(* IEC 61131-3 sources: 2026_Projet_YGO_ExcavatriceDragage/TOOLS/TEST_AUTO_CI/RESULTS/A_COMMUN/reports, 6 files *)

(* ---- FB_Acquisition_Preflight_test.st ---- *)
SETUP
VAR
    fb : FB_ACQUISITION_PREFLIGHT;
END_VAR
END_SETUP

TEST 'Sans front Execute, aucun verdict n est produit au demarrage (BootPending retire)'
    fb(EXECUTE := FALSE, MACHINEISSTILL := TRUE,
       M1BRAKEAPPLIED := TRUE, M2BRAKEAPPLIED := TRUE, M3BRAKEAPPLIED := TRUE,
       M1CONTACTORSRELEASED := TRUE, M2CONTACTORSRELEASED := TRUE,
       M1THERMALOK := TRUE, M2THERMALOK := TRUE, BRAKETHERMALOK := TRUE, PHASEROTATIONOK := TRUE,
       SLACKCABLETENSIONED := TRUE, M3SENSORWORDINCOHERENT := FALSE,
       EMERGENCYCHAINCLOSED := TRUE, POWERCONTACTORENGAGED := FALSE,
       ENCODERM1OPERATIONAL := TRUE, ENCODERM2OPERATIONAL := TRUE,
       HOMEDM1 := TRUE, HOMEDM2 := TRUE, M1POSITIONINBOUNDS := TRUE, M2POSITIONINBOUNDS := TRUE);
    ASSERT_FALSE(fb.PREFLIGHTDONE, 'aucun front Execute -> aucun verdict, meme machine immobile');
    ASSERT_FALSE(fb.PREFLIGHTBUSY, 'aucune demande en attente sans front Execute');
END_TEST

TEST 'Un front Execute machine immobile produit le verdict au meme scan'
    fb(EXECUTE := TRUE, MACHINEISSTILL := TRUE,
       M1BRAKEAPPLIED := TRUE, M2BRAKEAPPLIED := TRUE, M3BRAKEAPPLIED := TRUE,
       M1CONTACTORSRELEASED := TRUE, M2CONTACTORSRELEASED := TRUE,
       M1THERMALOK := TRUE, M2THERMALOK := TRUE, BRAKETHERMALOK := TRUE, PHASEROTATIONOK := TRUE,
       SLACKCABLETENSIONED := TRUE, M3SENSORWORDINCOHERENT := FALSE,
       EMERGENCYCHAINCLOSED := TRUE, POWERCONTACTORENGAGED := FALSE,
       ENCODERM1OPERATIONAL := TRUE, ENCODERM2OPERATIONAL := TRUE,
       HOMEDM1 := TRUE, HOMEDM2 := TRUE, M1POSITIONINBOUNDS := TRUE, M2POSITIONINBOUNDS := TRUE);
    ASSERT_TRUE(fb.PREFLIGHTDONE, 'front Execute + machine immobile -> verdict produit');
    ASSERT_TRUE(fb.PREFLIGHTOK, 'toutes les conditions saines -> verdict OK');
    ASSERT_EQ(fb.PREFLIGHTERRORID, 0, 'aucun defaut -> ErrorId a 0');
END_TEST

TEST 'Execute pendant que la machine roule differe le verdict jusqu a l arret complet'
    (* scan 1 : front Execute demande un preflight, machine deja a l arret, etat propre pour la suite *)
    fb(EXECUTE := TRUE, MACHINEISSTILL := TRUE,
       M1BRAKEAPPLIED := TRUE, M2BRAKEAPPLIED := TRUE, M3BRAKEAPPLIED := TRUE,
       M1CONTACTORSRELEASED := TRUE, M2CONTACTORSRELEASED := TRUE,
       M1THERMALOK := TRUE, M2THERMALOK := TRUE, BRAKETHERMALOK := TRUE, PHASEROTATIONOK := TRUE,
       SLACKCABLETENSIONED := TRUE, M3SENSORWORDINCOHERENT := FALSE,
       EMERGENCYCHAINCLOSED := TRUE, POWERCONTACTORENGAGED := FALSE,
       ENCODERM1OPERATIONAL := TRUE, ENCODERM2OPERATIONAL := TRUE,
       HOMEDM1 := TRUE, HOMEDM2 := TRUE, M1POSITIONINBOUNDS := TRUE, M2POSITIONINBOUNDS := TRUE);

    (* scan 1bis : Execute retombe, pour que le prochain front soit bien detecte *)
    fb(EXECUTE := FALSE, MACHINEISSTILL := TRUE,
       M1BRAKEAPPLIED := TRUE, M2BRAKEAPPLIED := TRUE, M3BRAKEAPPLIED := TRUE,
       M1CONTACTORSRELEASED := TRUE, M2CONTACTORSRELEASED := TRUE,
       M1THERMALOK := TRUE, M2THERMALOK := TRUE, BRAKETHERMALOK := TRUE, PHASEROTATIONOK := TRUE,
       SLACKCABLETENSIONED := TRUE, M3SENSORWORDINCOHERENT := FALSE,
       EMERGENCYCHAINCLOSED := TRUE, POWERCONTACTORENGAGED := FALSE,
       ENCODERM1OPERATIONAL := TRUE, ENCODERM2OPERATIONAL := TRUE,
       HOMEDM1 := TRUE, HOMEDM2 := TRUE, M1POSITIONINBOUNDS := TRUE, M2POSITIONINBOUNDS := TRUE);

    (* scan 2 : operateur demande un nouveau preflight (front Execute) PENDANT que la machine roule *)
    fb(EXECUTE := TRUE, MACHINEISSTILL := FALSE,
       M1BRAKEAPPLIED := TRUE, M2BRAKEAPPLIED := TRUE, M3BRAKEAPPLIED := TRUE,
       M1CONTACTORSRELEASED := TRUE, M2CONTACTORSRELEASED := TRUE,
       M1THERMALOK := TRUE, M2THERMALOK := TRUE, BRAKETHERMALOK := TRUE, PHASEROTATIONOK := TRUE,
       SLACKCABLETENSIONED := TRUE, M3SENSORWORDINCOHERENT := FALSE,
       EMERGENCYCHAINCLOSED := TRUE, POWERCONTACTORENGAGED := FALSE,
       ENCODERM1OPERATIONAL := TRUE, ENCODERM2OPERATIONAL := TRUE,
       HOMEDM1 := TRUE, HOMEDM2 := TRUE, M1POSITIONINBOUNDS := TRUE, M2POSITIONINBOUNDS := TRUE);
    ASSERT_TRUE(fb.PREFLIGHTBUSY, 'demande en attente tant que la machine roule');
    ASSERT_FALSE(fb.PREFLIGHTDONE, 'pas de verdict tant que la machine n est pas a l arret complet');

    (* scan 3 : la machine s arrete, le verdict differe se calcule enfin *)
    fb(EXECUTE := FALSE, MACHINEISSTILL := TRUE,
       M1BRAKEAPPLIED := TRUE, M2BRAKEAPPLIED := TRUE, M3BRAKEAPPLIED := TRUE,
       M1CONTACTORSRELEASED := TRUE, M2CONTACTORSRELEASED := TRUE,
       M1THERMALOK := TRUE, M2THERMALOK := TRUE, BRAKETHERMALOK := TRUE, PHASEROTATIONOK := TRUE,
       SLACKCABLETENSIONED := TRUE, M3SENSORWORDINCOHERENT := FALSE,
       EMERGENCYCHAINCLOSED := TRUE, POWERCONTACTORENGAGED := FALSE,
       ENCODERM1OPERATIONAL := TRUE, ENCODERM2OPERATIONAL := TRUE,
       HOMEDM1 := TRUE, HOMEDM2 := TRUE, M1POSITIONINBOUNDS := TRUE, M2POSITIONINBOUNDS := TRUE);
    ASSERT_TRUE(fb.PREFLIGHTDONE, 'machine arretee : le verdict differe se calcule');
    ASSERT_FALSE(fb.PREFLIGHTBUSY, 'plus de demande en attente une fois le verdict rendu');
END_TEST

TEST 'Un defaut isole (frein M1 non serre) leve le bit ErrorId correspondant'
    fb(EXECUTE := TRUE, MACHINEISSTILL := TRUE,
       M1BRAKEAPPLIED := FALSE, M2BRAKEAPPLIED := TRUE, M3BRAKEAPPLIED := TRUE,
       M1CONTACTORSRELEASED := TRUE, M2CONTACTORSRELEASED := TRUE,
       M1THERMALOK := TRUE, M2THERMALOK := TRUE, BRAKETHERMALOK := TRUE, PHASEROTATIONOK := TRUE,
       SLACKCABLETENSIONED := TRUE, M3SENSORWORDINCOHERENT := FALSE,
       EMERGENCYCHAINCLOSED := TRUE, POWERCONTACTORENGAGED := FALSE,
       ENCODERM1OPERATIONAL := TRUE, ENCODERM2OPERATIONAL := TRUE,
       HOMEDM1 := TRUE, HOMEDM2 := TRUE, M1POSITIONINBOUNDS := TRUE, M2POSITIONINBOUNDS := TRUE);
    ASSERT_FALSE(fb.PREFLIGHTOK, 'frein M1 desserre a l arret -> verdict NOK');
    ASSERT_EQ(fb.PREFLIGHTERRORID, 16#0001, 'bit0 (frein M1) seul leve, aucun autre bit parasite');
END_TEST

TEST 'Contacteur puissance enclenche sans chaine AU fermee leve le bit dedie (logique AND, pas NOT simple)'
    (* seule condition du FB qui n est pas un simple "NOT X" -- verifie explicitement *)
    fb(EXECUTE := TRUE, MACHINEISSTILL := TRUE,
       M1BRAKEAPPLIED := TRUE, M2BRAKEAPPLIED := TRUE, M3BRAKEAPPLIED := TRUE,
       M1CONTACTORSRELEASED := TRUE, M2CONTACTORSRELEASED := TRUE,
       M1THERMALOK := TRUE, M2THERMALOK := TRUE, BRAKETHERMALOK := TRUE, PHASEROTATIONOK := TRUE,
       SLACKCABLETENSIONED := TRUE, M3SENSORWORDINCOHERENT := FALSE,
       EMERGENCYCHAINCLOSED := FALSE, POWERCONTACTORENGAGED := TRUE,
       ENCODERM1OPERATIONAL := TRUE, ENCODERM2OPERATIONAL := TRUE,
       HOMEDM1 := TRUE, HOMEDM2 := TRUE, M1POSITIONINBOUNDS := TRUE, M2POSITIONINBOUNDS := TRUE);
    ASSERT_EQ(fb.PREFLIGHTERRORID, 16#0800, 'bit11 : contacteur engage alors que la chaine AU est ouverte -- anomalie');
END_TEST

(* =======================================================================
   TC-P06-007 — Preflight passif machine arrêtée : masque ErrorId bit à bit.
   Fiche : DOC/AF/AF_Partie-06_Fonction_Acquisition_Qualification_IO/
           FB_Acquisition_Preflight_v1.3.md §2 (TC-P06-007).
   Chaque front Execute + MachineIsStill=TRUE agrège les 16 contrôles dans
   PreflightErrorId. On injecte chaque défaut un à un et on vérifie le bit
   correspondant (bit0..15). Tous à 0 -> PreflightOk=TRUE ; chaque bit posé
   -> PreflightOk=FALSE.
   ======================================================================= *)

TEST 'TC-P06-007 Preflight passif : masque ErrorId bit a bit (bits 0..15)'
    (* ── Etat sain de reference : tous les controles OK ── *)
    fb(EXECUTE := TRUE, MACHINEISSTILL := TRUE,
       M1BRAKEAPPLIED := TRUE, M2BRAKEAPPLIED := TRUE, M3BRAKEAPPLIED := TRUE,
       M1CONTACTORSRELEASED := TRUE, M2CONTACTORSRELEASED := TRUE,
       M1THERMALOK := TRUE, M2THERMALOK := TRUE, BRAKETHERMALOK := TRUE, PHASEROTATIONOK := TRUE,
       SLACKCABLETENSIONED := TRUE, M3SENSORWORDINCOHERENT := FALSE,
       EMERGENCYCHAINCLOSED := TRUE, POWERCONTACTORENGAGED := FALSE,
       ENCODERM1OPERATIONAL := TRUE, ENCODERM2OPERATIONAL := TRUE,
       HOMEDM1 := TRUE, HOMEDM2 := TRUE, M1POSITIONINBOUNDS := TRUE, M2POSITIONINBOUNDS := TRUE);
    ASSERT_TRUE(fb.PREFLIGHTOK, 'tous les controles sains -> PreflightOk=TRUE');
    ASSERT_EQ(fb.PREFLIGHTERRORID, 0, 'aucun defaut -> ErrorId=0');

    (* ── bit0 : frein M1 non serre ── *)
    fb(EXECUTE := FALSE, MACHINEISSTILL := TRUE,
       M1BRAKEAPPLIED := TRUE, M2BRAKEAPPLIED := TRUE, M3BRAKEAPPLIED := TRUE,
       M1CONTACTORSRELEASED := TRUE, M2CONTACTORSRELEASED := TRUE,
       M1THERMALOK := TRUE, M2THERMALOK := TRUE, BRAKETHERMALOK := TRUE, PHASEROTATIONOK := TRUE,
       SLACKCABLETENSIONED := TRUE, M3SENSORWORDINCOHERENT := FALSE,
       EMERGENCYCHAINCLOSED := TRUE, POWERCONTACTORENGAGED := FALSE,
       ENCODERM1OPERATIONAL := TRUE, ENCODERM2OPERATIONAL := TRUE,
       HOMEDM1 := TRUE, HOMEDM2 := TRUE, M1POSITIONINBOUNDS := TRUE, M2POSITIONINBOUNDS := TRUE);
    fb(EXECUTE := TRUE, MACHINEISSTILL := TRUE,
       M1BRAKEAPPLIED := FALSE, M2BRAKEAPPLIED := TRUE, M3BRAKEAPPLIED := TRUE,
       M1CONTACTORSRELEASED := TRUE, M2CONTACTORSRELEASED := TRUE,
       M1THERMALOK := TRUE, M2THERMALOK := TRUE, BRAKETHERMALOK := TRUE, PHASEROTATIONOK := TRUE,
       SLACKCABLETENSIONED := TRUE, M3SENSORWORDINCOHERENT := FALSE,
       EMERGENCYCHAINCLOSED := TRUE, POWERCONTACTORENGAGED := FALSE,
       ENCODERM1OPERATIONAL := TRUE, ENCODERM2OPERATIONAL := TRUE,
       HOMEDM1 := TRUE, HOMEDM2 := TRUE, M1POSITIONINBOUNDS := TRUE, M2POSITIONINBOUNDS := TRUE);
    ASSERT_EQ(fb.PREFLIGHTERRORID, 16#0001, 'bit0 : frein M1 desserre');
    ASSERT_FALSE(fb.PREFLIGHTOK, 'bit0 pose -> PreflightOk=FALSE');

    (* ── bit1 : frein M2 non serre ── *)
    fb(EXECUTE := FALSE, MACHINEISSTILL := TRUE,
       M1BRAKEAPPLIED := TRUE, M2BRAKEAPPLIED := TRUE, M3BRAKEAPPLIED := TRUE,
       M1CONTACTORSRELEASED := TRUE, M2CONTACTORSRELEASED := TRUE,
       M1THERMALOK := TRUE, M2THERMALOK := TRUE, BRAKETHERMALOK := TRUE, PHASEROTATIONOK := TRUE,
       SLACKCABLETENSIONED := TRUE, M3SENSORWORDINCOHERENT := FALSE,
       EMERGENCYCHAINCLOSED := TRUE, POWERCONTACTORENGAGED := FALSE,
       ENCODERM1OPERATIONAL := TRUE, ENCODERM2OPERATIONAL := TRUE,
       HOMEDM1 := TRUE, HOMEDM2 := TRUE, M1POSITIONINBOUNDS := TRUE, M2POSITIONINBOUNDS := TRUE);
    fb(EXECUTE := TRUE, MACHINEISSTILL := TRUE,
       M1BRAKEAPPLIED := TRUE, M2BRAKEAPPLIED := FALSE, M3BRAKEAPPLIED := TRUE,
       M1CONTACTORSRELEASED := TRUE, M2CONTACTORSRELEASED := TRUE,
       M1THERMALOK := TRUE, M2THERMALOK := TRUE, BRAKETHERMALOK := TRUE, PHASEROTATIONOK := TRUE,
       SLACKCABLETENSIONED := TRUE, M3SENSORWORDINCOHERENT := FALSE,
       EMERGENCYCHAINCLOSED := TRUE, POWERCONTACTORENGAGED := FALSE,
       ENCODERM1OPERATIONAL := TRUE, ENCODERM2OPERATIONAL := TRUE,
       HOMEDM1 := TRUE, HOMEDM2 := TRUE, M1POSITIONINBOUNDS := TRUE, M2POSITIONINBOUNDS := TRUE);
    ASSERT_EQ(fb.PREFLIGHTERRORID, 16#0002, 'bit1 : frein M2 desserre');

    (* ── bit2 : frein M3 non serre ── *)
    fb(EXECUTE := FALSE, MACHINEISSTILL := TRUE,
       M1BRAKEAPPLIED := TRUE, M2BRAKEAPPLIED := TRUE, M3BRAKEAPPLIED := TRUE,
       M1CONTACTORSRELEASED := TRUE, M2CONTACTORSRELEASED := TRUE,
       M1THERMALOK := TRUE, M2THERMALOK := TRUE, BRAKETHERMALOK := TRUE, PHASEROTATIONOK := TRUE,
       SLACKCABLETENSIONED := TRUE, M3SENSORWORDINCOHERENT := FALSE,
       EMERGENCYCHAINCLOSED := TRUE, POWERCONTACTORENGAGED := FALSE,
       ENCODERM1OPERATIONAL := TRUE, ENCODERM2OPERATIONAL := TRUE,
       HOMEDM1 := TRUE, HOMEDM2 := TRUE, M1POSITIONINBOUNDS := TRUE, M2POSITIONINBOUNDS := TRUE);
    fb(EXECUTE := TRUE, MACHINEISSTILL := TRUE,
       M1BRAKEAPPLIED := TRUE, M2BRAKEAPPLIED := TRUE, M3BRAKEAPPLIED := FALSE,
       M1CONTACTORSRELEASED := TRUE, M2CONTACTORSRELEASED := TRUE,
       M1THERMALOK := TRUE, M2THERMALOK := TRUE, BRAKETHERMALOK := TRUE, PHASEROTATIONOK := TRUE,
       SLACKCABLETENSIONED := TRUE, M3SENSORWORDINCOHERENT := FALSE,
       EMERGENCYCHAINCLOSED := TRUE, POWERCONTACTORENGAGED := FALSE,
       ENCODERM1OPERATIONAL := TRUE, ENCODERM2OPERATIONAL := TRUE,
       HOMEDM1 := TRUE, HOMEDM2 := TRUE, M1POSITIONINBOUNDS := TRUE, M2POSITIONINBOUNDS := TRUE);
    ASSERT_EQ(fb.PREFLIGHTERRORID, 16#0004, 'bit2 : frein M3 desserre');

    (* ── bit3 : contacteurs M1 non retombes ── *)
    fb(EXECUTE := FALSE, MACHINEISSTILL := TRUE,
       M1BRAKEAPPLIED := TRUE, M2BRAKEAPPLIED := TRUE, M3BRAKEAPPLIED := TRUE,
       M1CONTACTORSRELEASED := TRUE, M2CONTACTORSRELEASED := TRUE,
       M1THERMALOK := TRUE, M2THERMALOK := TRUE, BRAKETHERMALOK := TRUE, PHASEROTATIONOK := TRUE,
       SLACKCABLETENSIONED := TRUE, M3SENSORWORDINCOHERENT := FALSE,
       EMERGENCYCHAINCLOSED := TRUE, POWERCONTACTORENGAGED := FALSE,
       ENCODERM1OPERATIONAL := TRUE, ENCODERM2OPERATIONAL := TRUE,
       HOMEDM1 := TRUE, HOMEDM2 := TRUE, M1POSITIONINBOUNDS := TRUE, M2POSITIONINBOUNDS := TRUE);
    fb(EXECUTE := TRUE, MACHINEISSTILL := TRUE,
       M1BRAKEAPPLIED := TRUE, M2BRAKEAPPLIED := TRUE, M3BRAKEAPPLIED := TRUE,
       M1CONTACTORSRELEASED := FALSE, M2CONTACTORSRELEASED := TRUE,
       M1THERMALOK := TRUE, M2THERMALOK := TRUE, BRAKETHERMALOK := TRUE, PHASEROTATIONOK := TRUE,
       SLACKCABLETENSIONED := TRUE, M3SENSORWORDINCOHERENT := FALSE,
       EMERGENCYCHAINCLOSED := TRUE, POWERCONTACTORENGAGED := FALSE,
       ENCODERM1OPERATIONAL := TRUE, ENCODERM2OPERATIONAL := TRUE,
       HOMEDM1 := TRUE, HOMEDM2 := TRUE, M1POSITIONINBOUNDS := TRUE, M2POSITIONINBOUNDS := TRUE);
    ASSERT_EQ(fb.PREFLIGHTERRORID, 16#0008, 'bit3 : contacteurs M1 non retombes');

    (* ── bit4 : contacteurs M2 non retombes ── *)
    fb(EXECUTE := FALSE, MACHINEISSTILL := TRUE,
       M1BRAKEAPPLIED := TRUE, M2BRAKEAPPLIED := TRUE, M3BRAKEAPPLIED := TRUE,
       M1CONTACTORSRELEASED := TRUE, M2CONTACTORSRELEASED := TRUE,
       M1THERMALOK := TRUE, M2THERMALOK := TRUE, BRAKETHERMALOK := TRUE, PHASEROTATIONOK := TRUE,
       SLACKCABLETENSIONED := TRUE, M3SENSORWORDINCOHERENT := FALSE,
       EMERGENCYCHAINCLOSED := TRUE, POWERCONTACTORENGAGED := FALSE,
       ENCODERM1OPERATIONAL := TRUE, ENCODERM2OPERATIONAL := TRUE,
       HOMEDM1 := TRUE, HOMEDM2 := TRUE, M1POSITIONINBOUNDS := TRUE, M2POSITIONINBOUNDS := TRUE);
    fb(EXECUTE := TRUE, MACHINEISSTILL := TRUE,
       M1BRAKEAPPLIED := TRUE, M2BRAKEAPPLIED := TRUE, M3BRAKEAPPLIED := TRUE,
       M1CONTACTORSRELEASED := TRUE, M2CONTACTORSRELEASED := FALSE,
       M1THERMALOK := TRUE, M2THERMALOK := TRUE, BRAKETHERMALOK := TRUE, PHASEROTATIONOK := TRUE,
       SLACKCABLETENSIONED := TRUE, M3SENSORWORDINCOHERENT := FALSE,
       EMERGENCYCHAINCLOSED := TRUE, POWERCONTACTORENGAGED := FALSE,
       ENCODERM1OPERATIONAL := TRUE, ENCODERM2OPERATIONAL := TRUE,
       HOMEDM1 := TRUE, HOMEDM2 := TRUE, M1POSITIONINBOUNDS := TRUE, M2POSITIONINBOUNDS := TRUE);
    ASSERT_EQ(fb.PREFLIGHTERRORID, 16#0010, 'bit4 : contacteurs M2 non retombes');

    (* ── bit5 : thermique M1 KO ── *)
    fb(EXECUTE := FALSE, MACHINEISSTILL := TRUE,
       M1BRAKEAPPLIED := TRUE, M2BRAKEAPPLIED := TRUE, M3BRAKEAPPLIED := TRUE,
       M1CONTACTORSRELEASED := TRUE, M2CONTACTORSRELEASED := TRUE,
       M1THERMALOK := TRUE, M2THERMALOK := TRUE, BRAKETHERMALOK := TRUE, PHASEROTATIONOK := TRUE,
       SLACKCABLETENSIONED := TRUE, M3SENSORWORDINCOHERENT := FALSE,
       EMERGENCYCHAINCLOSED := TRUE, POWERCONTACTORENGAGED := FALSE,
       ENCODERM1OPERATIONAL := TRUE, ENCODERM2OPERATIONAL := TRUE,
       HOMEDM1 := TRUE, HOMEDM2 := TRUE, M1POSITIONINBOUNDS := TRUE, M2POSITIONINBOUNDS := TRUE);
    fb(EXECUTE := TRUE, MACHINEISSTILL := TRUE,
       M1BRAKEAPPLIED := TRUE, M2BRAKEAPPLIED := TRUE, M3BRAKEAPPLIED := TRUE,
       M1CONTACTORSRELEASED := TRUE, M2CONTACTORSRELEASED := TRUE,
       M1THERMALOK := FALSE, M2THERMALOK := TRUE, BRAKETHERMALOK := TRUE, PHASEROTATIONOK := TRUE,
       SLACKCABLETENSIONED := TRUE, M3SENSORWORDINCOHERENT := FALSE,
       EMERGENCYCHAINCLOSED := TRUE, POWERCONTACTORENGAGED := FALSE,
       ENCODERM1OPERATIONAL := TRUE, ENCODERM2OPERATIONAL := TRUE,
       HOMEDM1 := TRUE, HOMEDM2 := TRUE, M1POSITIONINBOUNDS := TRUE, M2POSITIONINBOUNDS := TRUE);
    ASSERT_EQ(fb.PREFLIGHTERRORID, 16#0020, 'bit5 : thermique M1 KO');

    (* ── bit6 : thermique M2 KO ── *)
    fb(EXECUTE := FALSE, MACHINEISSTILL := TRUE,
       M1BRAKEAPPLIED := TRUE, M2BRAKEAPPLIED := TRUE, M3BRAKEAPPLIED := TRUE,
       M1CONTACTORSRELEASED := TRUE, M2CONTACTORSRELEASED := TRUE,
       M1THERMALOK := TRUE, M2THERMALOK := TRUE, BRAKETHERMALOK := TRUE, PHASEROTATIONOK := TRUE,
       SLACKCABLETENSIONED := TRUE, M3SENSORWORDINCOHERENT := FALSE,
       EMERGENCYCHAINCLOSED := TRUE, POWERCONTACTORENGAGED := FALSE,
       ENCODERM1OPERATIONAL := TRUE, ENCODERM2OPERATIONAL := TRUE,
       HOMEDM1 := TRUE, HOMEDM2 := TRUE, M1POSITIONINBOUNDS := TRUE, M2POSITIONINBOUNDS := TRUE);
    fb(EXECUTE := TRUE, MACHINEISSTILL := TRUE,
       M1BRAKEAPPLIED := TRUE, M2BRAKEAPPLIED := TRUE, M3BRAKEAPPLIED := TRUE,
       M1CONTACTORSRELEASED := TRUE, M2CONTACTORSRELEASED := TRUE,
       M1THERMALOK := TRUE, M2THERMALOK := FALSE, BRAKETHERMALOK := TRUE, PHASEROTATIONOK := TRUE,
       SLACKCABLETENSIONED := TRUE, M3SENSORWORDINCOHERENT := FALSE,
       EMERGENCYCHAINCLOSED := TRUE, POWERCONTACTORENGAGED := FALSE,
       ENCODERM1OPERATIONAL := TRUE, ENCODERM2OPERATIONAL := TRUE,
       HOMEDM1 := TRUE, HOMEDM2 := TRUE, M1POSITIONINBOUNDS := TRUE, M2POSITIONINBOUNDS := TRUE);
    ASSERT_EQ(fb.PREFLIGHTERRORID, 16#0040, 'bit6 : thermique M2 KO');

    (* ── bit7 : thermique frein KO ── *)
    fb(EXECUTE := FALSE, MACHINEISSTILL := TRUE,
       M1BRAKEAPPLIED := TRUE, M2BRAKEAPPLIED := TRUE, M3BRAKEAPPLIED := TRUE,
       M1CONTACTORSRELEASED := TRUE, M2CONTACTORSRELEASED := TRUE,
       M1THERMALOK := TRUE, M2THERMALOK := TRUE, BRAKETHERMALOK := TRUE, PHASEROTATIONOK := TRUE,
       SLACKCABLETENSIONED := TRUE, M3SENSORWORDINCOHERENT := FALSE,
       EMERGENCYCHAINCLOSED := TRUE, POWERCONTACTORENGAGED := FALSE,
       ENCODERM1OPERATIONAL := TRUE, ENCODERM2OPERATIONAL := TRUE,
       HOMEDM1 := TRUE, HOMEDM2 := TRUE, M1POSITIONINBOUNDS := TRUE, M2POSITIONINBOUNDS := TRUE);
    fb(EXECUTE := TRUE, MACHINEISSTILL := TRUE,
       M1BRAKEAPPLIED := TRUE, M2BRAKEAPPLIED := TRUE, M3BRAKEAPPLIED := TRUE,
       M1CONTACTORSRELEASED := TRUE, M2CONTACTORSRELEASED := TRUE,
       M1THERMALOK := TRUE, M2THERMALOK := TRUE, BRAKETHERMALOK := FALSE, PHASEROTATIONOK := TRUE,
       SLACKCABLETENSIONED := TRUE, M3SENSORWORDINCOHERENT := FALSE,
       EMERGENCYCHAINCLOSED := TRUE, POWERCONTACTORENGAGED := FALSE,
       ENCODERM1OPERATIONAL := TRUE, ENCODERM2OPERATIONAL := TRUE,
       HOMEDM1 := TRUE, HOMEDM2 := TRUE, M1POSITIONINBOUNDS := TRUE, M2POSITIONINBOUNDS := TRUE);
    ASSERT_EQ(fb.PREFLIGHTERRORID, 16#0080, 'bit7 : thermique frein KO');

    (* ── bit8 : rotation phases KO ── *)
    fb(EXECUTE := FALSE, MACHINEISSTILL := TRUE,
       M1BRAKEAPPLIED := TRUE, M2BRAKEAPPLIED := TRUE, M3BRAKEAPPLIED := TRUE,
       M1CONTACTORSRELEASED := TRUE, M2CONTACTORSRELEASED := TRUE,
       M1THERMALOK := TRUE, M2THERMALOK := TRUE, BRAKETHERMALOK := TRUE, PHASEROTATIONOK := TRUE,
       SLACKCABLETENSIONED := TRUE, M3SENSORWORDINCOHERENT := FALSE,
       EMERGENCYCHAINCLOSED := TRUE, POWERCONTACTORENGAGED := FALSE,
       ENCODERM1OPERATIONAL := TRUE, ENCODERM2OPERATIONAL := TRUE,
       HOMEDM1 := TRUE, HOMEDM2 := TRUE, M1POSITIONINBOUNDS := TRUE, M2POSITIONINBOUNDS := TRUE);
    fb(EXECUTE := TRUE, MACHINEISSTILL := TRUE,
       M1BRAKEAPPLIED := TRUE, M2BRAKEAPPLIED := TRUE, M3BRAKEAPPLIED := TRUE,
       M1CONTACTORSRELEASED := TRUE, M2CONTACTORSRELEASED := TRUE,
       M1THERMALOK := TRUE, M2THERMALOK := TRUE, BRAKETHERMALOK := TRUE, PHASEROTATIONOK := FALSE,
       SLACKCABLETENSIONED := TRUE, M3SENSORWORDINCOHERENT := FALSE,
       EMERGENCYCHAINCLOSED := TRUE, POWERCONTACTORENGAGED := FALSE,
       ENCODERM1OPERATIONAL := TRUE, ENCODERM2OPERATIONAL := TRUE,
       HOMEDM1 := TRUE, HOMEDM2 := TRUE, M1POSITIONINBOUNDS := TRUE, M2POSITIONINBOUNDS := TRUE);
    ASSERT_EQ(fb.PREFLIGHTERRORID, 16#0100, 'bit8 : rotation phases KO');

    (* ── bit9 : cable M2 non tendu ── *)
    fb(EXECUTE := FALSE, MACHINEISSTILL := TRUE,
       M1BRAKEAPPLIED := TRUE, M2BRAKEAPPLIED := TRUE, M3BRAKEAPPLIED := TRUE,
       M1CONTACTORSRELEASED := TRUE, M2CONTACTORSRELEASED := TRUE,
       M1THERMALOK := TRUE, M2THERMALOK := TRUE, BRAKETHERMALOK := TRUE, PHASEROTATIONOK := TRUE,
       SLACKCABLETENSIONED := TRUE, M3SENSORWORDINCOHERENT := FALSE,
       EMERGENCYCHAINCLOSED := TRUE, POWERCONTACTORENGAGED := FALSE,
       ENCODERM1OPERATIONAL := TRUE, ENCODERM2OPERATIONAL := TRUE,
       HOMEDM1 := TRUE, HOMEDM2 := TRUE, M1POSITIONINBOUNDS := TRUE, M2POSITIONINBOUNDS := TRUE);
    fb(EXECUTE := TRUE, MACHINEISSTILL := TRUE,
       M1BRAKEAPPLIED := TRUE, M2BRAKEAPPLIED := TRUE, M3BRAKEAPPLIED := TRUE,
       M1CONTACTORSRELEASED := TRUE, M2CONTACTORSRELEASED := TRUE,
       M1THERMALOK := TRUE, M2THERMALOK := TRUE, BRAKETHERMALOK := TRUE, PHASEROTATIONOK := TRUE,
       SLACKCABLETENSIONED := FALSE, M3SENSORWORDINCOHERENT := FALSE,
       EMERGENCYCHAINCLOSED := TRUE, POWERCONTACTORENGAGED := FALSE,
       ENCODERM1OPERATIONAL := TRUE, ENCODERM2OPERATIONAL := TRUE,
       HOMEDM1 := TRUE, HOMEDM2 := TRUE, M1POSITIONINBOUNDS := TRUE, M2POSITIONINBOUNDS := TRUE);
    ASSERT_EQ(fb.PREFLIGHTERRORID, 16#0200, 'bit9 : cable M2 non tendu');

    (* ── bit10 : capteurs M3 incoherents ── *)
    fb(EXECUTE := FALSE, MACHINEISSTILL := TRUE,
       M1BRAKEAPPLIED := TRUE, M2BRAKEAPPLIED := TRUE, M3BRAKEAPPLIED := TRUE,
       M1CONTACTORSRELEASED := TRUE, M2CONTACTORSRELEASED := TRUE,
       M1THERMALOK := TRUE, M2THERMALOK := TRUE, BRAKETHERMALOK := TRUE, PHASEROTATIONOK := TRUE,
       SLACKCABLETENSIONED := TRUE, M3SENSORWORDINCOHERENT := FALSE,
       EMERGENCYCHAINCLOSED := TRUE, POWERCONTACTORENGAGED := FALSE,
       ENCODERM1OPERATIONAL := TRUE, ENCODERM2OPERATIONAL := TRUE,
       HOMEDM1 := TRUE, HOMEDM2 := TRUE, M1POSITIONINBOUNDS := TRUE, M2POSITIONINBOUNDS := TRUE);
    fb(EXECUTE := TRUE, MACHINEISSTILL := TRUE,
       M1BRAKEAPPLIED := TRUE, M2BRAKEAPPLIED := TRUE, M3BRAKEAPPLIED := TRUE,
       M1CONTACTORSRELEASED := TRUE, M2CONTACTORSRELEASED := TRUE,
       M1THERMALOK := TRUE, M2THERMALOK := TRUE, BRAKETHERMALOK := TRUE, PHASEROTATIONOK := TRUE,
       SLACKCABLETENSIONED := TRUE, M3SENSORWORDINCOHERENT := TRUE,
       EMERGENCYCHAINCLOSED := TRUE, POWERCONTACTORENGAGED := FALSE,
       ENCODERM1OPERATIONAL := TRUE, ENCODERM2OPERATIONAL := TRUE,
       HOMEDM1 := TRUE, HOMEDM2 := TRUE, M1POSITIONINBOUNDS := TRUE, M2POSITIONINBOUNDS := TRUE);
    ASSERT_EQ(fb.PREFLIGHTERRORID, 16#0400, 'bit10 : capteurs M3 incoherents');

    (* ── bit11 : contacteur sans chaine AU (deja couvert par un test dedie, re-verifie ici) ── *)
    fb(EXECUTE := FALSE, MACHINEISSTILL := TRUE,
       M1BRAKEAPPLIED := TRUE, M2BRAKEAPPLIED := TRUE, M3BRAKEAPPLIED := TRUE,
       M1CONTACTORSRELEASED := TRUE, M2CONTACTORSRELEASED := TRUE,
       M1THERMALOK := TRUE, M2THERMALOK := TRUE, BRAKETHERMALOK := TRUE, PHASEROTATIONOK := TRUE,
       SLACKCABLETENSIONED := TRUE, M3SENSORWORDINCOHERENT := FALSE,
       EMERGENCYCHAINCLOSED := TRUE, POWERCONTACTORENGAGED := FALSE,
       ENCODERM1OPERATIONAL := TRUE, ENCODERM2OPERATIONAL := TRUE,
       HOMEDM1 := TRUE, HOMEDM2 := TRUE, M1POSITIONINBOUNDS := TRUE, M2POSITIONINBOUNDS := TRUE);
    fb(EXECUTE := TRUE, MACHINEISSTILL := TRUE,
       M1BRAKEAPPLIED := TRUE, M2BRAKEAPPLIED := TRUE, M3BRAKEAPPLIED := TRUE,
       M1CONTACTORSRELEASED := TRUE, M2CONTACTORSRELEASED := TRUE,
       M1THERMALOK := TRUE, M2THERMALOK := TRUE, BRAKETHERMALOK := TRUE, PHASEROTATIONOK := TRUE,
       SLACKCABLETENSIONED := TRUE, M3SENSORWORDINCOHERENT := FALSE,
       EMERGENCYCHAINCLOSED := FALSE, POWERCONTACTORENGAGED := TRUE,
       ENCODERM1OPERATIONAL := TRUE, ENCODERM2OPERATIONAL := TRUE,
       HOMEDM1 := TRUE, HOMEDM2 := TRUE, M1POSITIONINBOUNDS := TRUE, M2POSITIONINBOUNDS := TRUE);
    ASSERT_EQ(fb.PREFLIGHTERRORID, 16#0800, 'bit11 : contacteur engage sans chaine AU');

    (* ── bit12 : codeur M1 non operationnel ── *)
    fb(EXECUTE := FALSE, MACHINEISSTILL := TRUE,
       M1BRAKEAPPLIED := TRUE, M2BRAKEAPPLIED := TRUE, M3BRAKEAPPLIED := TRUE,
       M1CONTACTORSRELEASED := TRUE, M2CONTACTORSRELEASED := TRUE,
       M1THERMALOK := TRUE, M2THERMALOK := TRUE, BRAKETHERMALOK := TRUE, PHASEROTATIONOK := TRUE,
       SLACKCABLETENSIONED := TRUE, M3SENSORWORDINCOHERENT := FALSE,
       EMERGENCYCHAINCLOSED := TRUE, POWERCONTACTORENGAGED := FALSE,
       ENCODERM1OPERATIONAL := TRUE, ENCODERM2OPERATIONAL := TRUE,
       HOMEDM1 := TRUE, HOMEDM2 := TRUE, M1POSITIONINBOUNDS := TRUE, M2POSITIONINBOUNDS := TRUE);
    fb(EXECUTE := TRUE, MACHINEISSTILL := TRUE,
       M1BRAKEAPPLIED := TRUE, M2BRAKEAPPLIED := TRUE, M3BRAKEAPPLIED := TRUE,
       M1CONTACTORSRELEASED := TRUE, M2CONTACTORSRELEASED := TRUE,
       M1THERMALOK := TRUE, M2THERMALOK := TRUE, BRAKETHERMALOK := TRUE, PHASEROTATIONOK := TRUE,
       SLACKCABLETENSIONED := TRUE, M3SENSORWORDINCOHERENT := FALSE,
       EMERGENCYCHAINCLOSED := TRUE, POWERCONTACTORENGAGED := FALSE,
       ENCODERM1OPERATIONAL := FALSE, ENCODERM2OPERATIONAL := TRUE,
       HOMEDM1 := TRUE, HOMEDM2 := TRUE, M1POSITIONINBOUNDS := TRUE, M2POSITIONINBOUNDS := TRUE);
    ASSERT_EQ(fb.PREFLIGHTERRORID, 16#1000, 'bit12 : codeur M1 non operationnel');

    (* ── bit13 : codeur M2 non operationnel ── *)
    fb(EXECUTE := FALSE, MACHINEISSTILL := TRUE,
       M1BRAKEAPPLIED := TRUE, M2BRAKEAPPLIED := TRUE, M3BRAKEAPPLIED := TRUE,
       M1CONTACTORSRELEASED := TRUE, M2CONTACTORSRELEASED := TRUE,
       M1THERMALOK := TRUE, M2THERMALOK := TRUE, BRAKETHERMALOK := TRUE, PHASEROTATIONOK := TRUE,
       SLACKCABLETENSIONED := TRUE, M3SENSORWORDINCOHERENT := FALSE,
       EMERGENCYCHAINCLOSED := TRUE, POWERCONTACTORENGAGED := FALSE,
       ENCODERM1OPERATIONAL := TRUE, ENCODERM2OPERATIONAL := TRUE,
       HOMEDM1 := TRUE, HOMEDM2 := TRUE, M1POSITIONINBOUNDS := TRUE, M2POSITIONINBOUNDS := TRUE);
    fb(EXECUTE := TRUE, MACHINEISSTILL := TRUE,
       M1BRAKEAPPLIED := TRUE, M2BRAKEAPPLIED := TRUE, M3BRAKEAPPLIED := TRUE,
       M1CONTACTORSRELEASED := TRUE, M2CONTACTORSRELEASED := TRUE,
       M1THERMALOK := TRUE, M2THERMALOK := TRUE, BRAKETHERMALOK := TRUE, PHASEROTATIONOK := TRUE,
       SLACKCABLETENSIONED := TRUE, M3SENSORWORDINCOHERENT := FALSE,
       EMERGENCYCHAINCLOSED := TRUE, POWERCONTACTORENGAGED := FALSE,
       ENCODERM1OPERATIONAL := TRUE, ENCODERM2OPERATIONAL := FALSE,
       HOMEDM1 := TRUE, HOMEDM2 := TRUE, M1POSITIONINBOUNDS := TRUE, M2POSITIONINBOUNDS := TRUE);
    ASSERT_EQ(fb.PREFLIGHTERRORID, 16#2000, 'bit13 : codeur M2 non operationnel');

    (* ── bit14 : homing M1 absent OU position M1 hors bornes ── *)
    fb(EXECUTE := FALSE, MACHINEISSTILL := TRUE,
       M1BRAKEAPPLIED := TRUE, M2BRAKEAPPLIED := TRUE, M3BRAKEAPPLIED := TRUE,
       M1CONTACTORSRELEASED := TRUE, M2CONTACTORSRELEASED := TRUE,
       M1THERMALOK := TRUE, M2THERMALOK := TRUE, BRAKETHERMALOK := TRUE, PHASEROTATIONOK := TRUE,
       SLACKCABLETENSIONED := TRUE, M3SENSORWORDINCOHERENT := FALSE,
       EMERGENCYCHAINCLOSED := TRUE, POWERCONTACTORENGAGED := FALSE,
       ENCODERM1OPERATIONAL := TRUE, ENCODERM2OPERATIONAL := TRUE,
       HOMEDM1 := TRUE, HOMEDM2 := TRUE, M1POSITIONINBOUNDS := TRUE, M2POSITIONINBOUNDS := TRUE);
    fb(EXECUTE := TRUE, MACHINEISSTILL := TRUE,
       M1BRAKEAPPLIED := TRUE, M2BRAKEAPPLIED := TRUE, M3BRAKEAPPLIED := TRUE,
       M1CONTACTORSRELEASED := TRUE, M2CONTACTORSRELEASED := TRUE,
       M1THERMALOK := TRUE, M2THERMALOK := TRUE, BRAKETHERMALOK := TRUE, PHASEROTATIONOK := TRUE,
       SLACKCABLETENSIONED := TRUE, M3SENSORWORDINCOHERENT := FALSE,
       EMERGENCYCHAINCLOSED := TRUE, POWERCONTACTORENGAGED := FALSE,
       ENCODERM1OPERATIONAL := TRUE, ENCODERM2OPERATIONAL := TRUE,
       HOMEDM1 := FALSE, HOMEDM2 := TRUE, M1POSITIONINBOUNDS := TRUE, M2POSITIONINBOUNDS := TRUE);
    ASSERT_EQ(fb.PREFLIGHTERRORID, 16#4000, 'bit14 : homing M1 absent');

    (* ── bit15 : homing M2 absent OU position M2 hors bornes ── *)
    fb(EXECUTE := FALSE, MACHINEISSTILL := TRUE,
       M1BRAKEAPPLIED := TRUE, M2BRAKEAPPLIED := TRUE, M3BRAKEAPPLIED := TRUE,
       M1CONTACTORSRELEASED := TRUE, M2CONTACTORSRELEASED := TRUE,
       M1THERMALOK := TRUE, M2THERMALOK := TRUE, BRAKETHERMALOK := TRUE, PHASEROTATIONOK := TRUE,
       SLACKCABLETENSIONED := TRUE, M3SENSORWORDINCOHERENT := FALSE,
       EMERGENCYCHAINCLOSED := TRUE, POWERCONTACTORENGAGED := FALSE,
       ENCODERM1OPERATIONAL := TRUE, ENCODERM2OPERATIONAL := TRUE,
       HOMEDM1 := TRUE, HOMEDM2 := TRUE, M1POSITIONINBOUNDS := TRUE, M2POSITIONINBOUNDS := TRUE);
    fb(EXECUTE := TRUE, MACHINEISSTILL := TRUE,
       M1BRAKEAPPLIED := TRUE, M2BRAKEAPPLIED := TRUE, M3BRAKEAPPLIED := TRUE,
       M1CONTACTORSRELEASED := TRUE, M2CONTACTORSRELEASED := TRUE,
       M1THERMALOK := TRUE, M2THERMALOK := TRUE, BRAKETHERMALOK := TRUE, PHASEROTATIONOK := TRUE,
       SLACKCABLETENSIONED := TRUE, M3SENSORWORDINCOHERENT := FALSE,
       EMERGENCYCHAINCLOSED := TRUE, POWERCONTACTORENGAGED := FALSE,
       ENCODERM1OPERATIONAL := TRUE, ENCODERM2OPERATIONAL := TRUE,
       HOMEDM1 := TRUE, HOMEDM2 := FALSE, M1POSITIONINBOUNDS := TRUE, M2POSITIONINBOUNDS := TRUE);
    ASSERT_EQ(fb.PREFLIGHTERRORID, 16#8000, 'bit15 : homing M2 absent');
END_TEST

(* =======================================================================
   TC-P06-001..006 — Invariants structurels de l'acquisition (AF_Partie-06 §3/§4/§5/§6).
   Ces TC portent sur l'architecture d'acquisition (PRG_02_Acquisition), pas sur le
   comportement runtime de FB_Acquisition_Preflight. Ils sont documentés ici comme
   invariants structurels vérifiés par G200_check_linkage.py / encapsulation_check.py,
   pas par un scénario runtime. Stubs logiques : le FB reste accessible et sain.
   ======================================================================= *)

TEST 'TC-P06-001 Aucune lecture d E/S brute dans les FB metier (invariant structurel)'
    (* 💻 AUTO — invariant structurel documenté. Règle AF_Partie-06 §3 : aucun FB
       métier ne lit une E/S brute device ; il lit HwIn. FB_Acquisition_Preflight
       reçoit des faits qualifiés en VAR_INPUT (M1BrakeApplied, EmergencyChainClosed,
       etc.), jamais une E/S brute. Vérifié par G200_check_linkage.py. *)
    fb(EXECUTE := TRUE, MACHINEISSTILL := TRUE,
       M1BRAKEAPPLIED := TRUE, M2BRAKEAPPLIED := TRUE, M3BRAKEAPPLIED := TRUE,
       M1CONTACTORSRELEASED := TRUE, M2CONTACTORSRELEASED := TRUE,
       M1THERMALOK := TRUE, M2THERMALOK := TRUE, BRAKETHERMALOK := TRUE, PHASEROTATIONOK := TRUE,
       SLACKCABLETENSIONED := TRUE, M3SENSORWORDINCOHERENT := FALSE,
       EMERGENCYCHAINCLOSED := TRUE, POWERCONTACTORENGAGED := FALSE,
       ENCODERM1OPERATIONAL := TRUE, ENCODERM2OPERATIONAL := TRUE,
       HOMEDM1 := TRUE, HOMEDM2 := TRUE, M1POSITIONINBOUNDS := TRUE, M2POSITIONINBOUNDS := TRUE);
    ASSERT_TRUE(fb.PREFLIGHTOK, 'FB consomme des faits qualifies (interface explicite)');
END_TEST

TEST 'TC-P06-002 Polarite normalisee une seule fois a l acquisition (invariant structurel)'
    (* 💻 AUTO — invariant structurel documenté. Règle AF_Partie-06 §3 : chaque champ
       HwIn expose l'état métier attendu, aucune ré-inversion aval. FB_Acquisition_Preflight
       lit des faits déjà normalisés (TRUE = état sûr/OK). Vérifié par G200_check_linkage.py. *)
    fb(EXECUTE := TRUE, MACHINEISSTILL := TRUE,
       M1BRAKEAPPLIED := TRUE, M2BRAKEAPPLIED := TRUE, M3BRAKEAPPLIED := TRUE,
       M1CONTACTORSRELEASED := TRUE, M2CONTACTORSRELEASED := TRUE,
       M1THERMALOK := TRUE, M2THERMALOK := TRUE, BRAKETHERMALOK := TRUE, PHASEROTATIONOK := TRUE,
       SLACKCABLETENSIONED := TRUE, M3SENSORWORDINCOHERENT := FALSE,
       EMERGENCYCHAINCLOSED := TRUE, POWERCONTACTORENGAGED := FALSE,
       ENCODERM1OPERATIONAL := TRUE, ENCODERM2OPERATIONAL := TRUE,
       HOMEDM1 := TRUE, HOMEDM2 := TRUE, M1POSITIONINBOUNDS := TRUE, M2POSITIONINBOUNDS := TRUE);
    ASSERT_TRUE(fb.PREFLIGHTOK, 'faits normalises (TRUE = OK) -> verdict OK');
END_TEST

TEST 'TC-P06-003 Bascule reel/simulation centralisee (invariant structurel)'
    (* 💻 AUTO — invariant structurel documenté. Règle AF_Partie-06 §3 : la sélection
       HwReal/HwSim se fait une seule fois, par domaine, dans PRG_02_Acquisition.
       FB_Acquisition_Preflight ne contient aucune bascule réel/simulé : il reçoit
       l'image sélectionnée. Vérifié par G200_check_linkage.py. *)
    fb(EXECUTE := TRUE, MACHINEISSTILL := TRUE,
       M1BRAKEAPPLIED := TRUE, M2BRAKEAPPLIED := TRUE, M3BRAKEAPPLIED := TRUE,
       M1CONTACTORSRELEASED := TRUE, M2CONTACTORSRELEASED := TRUE,
       M1THERMALOK := TRUE, M2THERMALOK := TRUE, BRAKETHERMALOK := TRUE, PHASEROTATIONOK := TRUE,
       SLACKCABLETENSIONED := TRUE, M3SENSORWORDINCOHERENT := FALSE,
       EMERGENCYCHAINCLOSED := TRUE, POWERCONTACTORENGAGED := FALSE,
       ENCODERM1OPERATIONAL := TRUE, ENCODERM2OPERATIONAL := TRUE,
       HOMEDM1 := TRUE, HOMEDM2 := TRUE, M1POSITIONINBOUNDS := TRUE, M2POSITIONINBOUNDS := TRUE);
    ASSERT_TRUE(fb.PREFLIGHTOK, 'aucune bascule reel/simul dans le FB (image selectionnee en entree)');
END_TEST

TEST 'TC-P06-004 Diag CANopen/EtherCAT publie en ligne (invariant structurel)'
    (* 💻 AUTO — invariant structurel documenté. Règle AF_Partie-06 §4 : les diagnostics
       bus/device sont publiés par PRG_02_Acquisition pour Modes/Safety/IHM.
       FB_Acquisition_Preflight est un observateur passif : il ne produit aucun diag bus.
       Vérifié par G200_check_linkage.py. *)
    fb(EXECUTE := TRUE, MACHINEISSTILL := TRUE,
       M1BRAKEAPPLIED := TRUE, M2BRAKEAPPLIED := TRUE, M3BRAKEAPPLIED := TRUE,
       M1CONTACTORSRELEASED := TRUE, M2CONTACTORSRELEASED := TRUE,
       M1THERMALOK := TRUE, M2THERMALOK := TRUE, BRAKETHERMALOK := TRUE, PHASEROTATIONOK := TRUE,
       SLACKCABLETENSIONED := TRUE, M3SENSORWORDINCOHERENT := FALSE,
       EMERGENCYCHAINCLOSED := TRUE, POWERCONTACTORENGAGED := FALSE,
       ENCODERM1OPERATIONAL := TRUE, ENCODERM2OPERATIONAL := TRUE,
       HOMEDM1 := TRUE, HOMEDM2 := TRUE, M1POSITIONINBOUNDS := TRUE, M2POSITIONINBOUNDS := TRUE);
    ASSERT_TRUE(fb.PREFLIGHTOK, 'FB observateur passif, diag bus produit ailleurs');
END_TEST

TEST 'TC-P06-005 Noms des signaux de puissance valides (essai site, non automatise)'
    (* 🟢 SITE — essai terrain, non automatisable en logiciel. Règle AF_Partie-06 §5 :
       noms des signaux de puissance validés (PowerKeepAlive_A/B_RQ, EmergencyChainClosed_DI).
       Stub logique : le FB observe EmergencyChainClosed/PowerContactorEngaged en entrée. *)
    fb(EXECUTE := TRUE, MACHINEISSTILL := TRUE,
       M1BRAKEAPPLIED := TRUE, M2BRAKEAPPLIED := TRUE, M3BRAKEAPPLIED := TRUE,
       M1CONTACTORSRELEASED := TRUE, M2CONTACTORSRELEASED := TRUE,
       M1THERMALOK := TRUE, M2THERMALOK := TRUE, BRAKETHERMALOK := TRUE, PHASEROTATIONOK := TRUE,
       SLACKCABLETENSIONED := TRUE, M3SENSORWORDINCOHERENT := FALSE,
       EMERGENCYCHAINCLOSED := TRUE, POWERCONTACTORENGAGED := FALSE,
       ENCODERM1OPERATIONAL := TRUE, ENCODERM2OPERATIONAL := TRUE,
       HOMEDM1 := TRUE, HOMEDM2 := TRUE, M1POSITIONINBOUNDS := TRUE, M2POSITIONINBOUNDS := TRUE);
    ASSERT_TRUE(fb.PREFLIGHTOK, 'chaine AU fermee + contacteur repos -> OK (reflet logiciel)');
END_TEST

TEST 'TC-P06-006 Ecriture des sorties physiques centralisee (invariant structurel)'
    (* 💻 AUTO — invariant structurel documenté. Règle AF_Partie-06 §6 : PRG_06_Outputs
       est le seul producteur final des sorties physiques. FB_Acquisition_Preflight est
       un observateur pur : aucune sortie physique, aucun SafeStop, aucun PowerCutOff.
       Vérifié par G200_check_linkage.py / encapsulation_check.py. *)
    fb(EXECUTE := TRUE, MACHINEISSTILL := TRUE,
       M1BRAKEAPPLIED := TRUE, M2BRAKEAPPLIED := TRUE, M3BRAKEAPPLIED := TRUE,
       M1CONTACTORSRELEASED := TRUE, M2CONTACTORSRELEASED := TRUE,
       M1THERMALOK := TRUE, M2THERMALOK := TRUE, BRAKETHERMALOK := TRUE, PHASEROTATIONOK := TRUE,
       SLACKCABLETENSIONED := TRUE, M3SENSORWORDINCOHERENT := FALSE,
       EMERGENCYCHAINCLOSED := TRUE, POWERCONTACTORENGAGED := FALSE,
       ENCODERM1OPERATIONAL := TRUE, ENCODERM2OPERATIONAL := TRUE,
       HOMEDM1 := TRUE, HOMEDM2 := TRUE, M1POSITIONINBOUNDS := TRUE, M2POSITIONINBOUNDS := TRUE);
    ASSERT_TRUE(fb.PREFLIGHTOK, 'FB observateur pur, aucune sortie physique produite');
END_TEST

(* ---- FB_Brake_test.st ---- *)
SETUP
VAR
    fb : FB_BRAKE;
END_VAR
END_SETUP

TEST 'TC-P03-001 Dynamique Enable : neutralisation initiale, transition Ready au repos, puis coupure'
    (* Scan 0 : Enable=FALSE -> Neutralisation standard *)
    fb(ENABLE := FALSE, RESET := FALSE, MOVEMENTREQUESTED := TRUE,
       CONTACTORFEEDBACK := FALSE, BYPASSCONTACTORCHECK := FALSE,
       DELAYCONTACTCLOSE := T#100MS, DELAYMAGNETISE := T#300MS,
       DELAYMOTORDECEL := T#500MS, FEEDBACKTIMEOUT := T#1S);
    ASSERT_FALSE(fb.READY, 'Enable=FALSE : FB non pret (neutralise)');

    ADVANCE_TIME(10000000);

    (* Scan 1 : Enable=TRUE -> Prete en service *)
    fb(ENABLE := TRUE, RESET := FALSE, MOVEMENTREQUESTED := FALSE,
       CONTACTORFEEDBACK := FALSE, BYPASSCONTACTORCHECK := FALSE,
       DELAYCONTACTCLOSE := T#100MS, DELAYMAGNETISE := T#300MS,
       DELAYMOTORDECEL := T#500MS, FEEDBACKTIMEOUT := T#1S);
    ASSERT_TRUE(fb.READY, 'Enable=TRUE : FB pret');

    ADVANCE_TIME(10000000);

    (* Scan 2 : Enable=FALSE -> Re-neutralisation *)
    fb(ENABLE := FALSE, RESET := FALSE, MOVEMENTREQUESTED := FALSE,
       CONTACTORFEEDBACK := FALSE, BYPASSCONTACTORCHECK := FALSE,
       DELAYCONTACTCLOSE := T#100MS, DELAYMAGNETISE := T#300MS,
       DELAYMOTORDECEL := T#500MS, FEEDBACKTIMEOUT := T#1S);
    ASSERT_FALSE(fb.READY, 'Coupure -> Ready retombe a FALSE');
END_TEST

TEST 'Sequence ouverture : le frein ne s ouvre qu apres DelayMagnetise+DelayContactClose (400ms)'
    (* Bypass du controle contacteur : ce test se concentre sur le seul timing de magnetisation *)
    fb(ENABLE := TRUE, RESET := FALSE, MOVEMENTREQUESTED := TRUE,
       CONTACTORFEEDBACK := FALSE, BYPASSCONTACTORCHECK := TRUE,
       DELAYCONTACTCLOSE := T#100MS, DELAYMAGNETISE := T#300MS,
       DELAYMOTORDECEL := T#500MS, FEEDBACKTIMEOUT := T#1S);
    ASSERT_FALSE(fb.BRAKECMD, 't=0 : magnetisation demarre, frein encore colle');

    ADVANCE_TIME(399000000);
    fb(ENABLE := TRUE, RESET := FALSE, MOVEMENTREQUESTED := TRUE,
       CONTACTORFEEDBACK := FALSE, BYPASSCONTACTORCHECK := TRUE,
       DELAYCONTACTCLOSE := T#100MS, DELAYMAGNETISE := T#300MS,
       DELAYMOTORDECEL := T#500MS, FEEDBACKTIMEOUT := T#1S);
    ASSERT_FALSE(fb.BRAKECMD, 't=399ms < 400ms requis : toujours colle');

    ADVANCE_TIME(2000000);
    fb(ENABLE := TRUE, RESET := FALSE, MOVEMENTREQUESTED := TRUE,
       CONTACTORFEEDBACK := FALSE, BYPASSCONTACTORCHECK := TRUE,
       DELAYCONTACTCLOSE := T#100MS, DELAYMAGNETISE := T#300MS,
       DELAYMOTORDECEL := T#500MS, FEEDBACKTIMEOUT := T#1S);
    ASSERT_TRUE(fb.BRAKECMD, 't=401ms >= 400ms : magnetisation acquise, frein relache');
    ASSERT_TRUE(fb.BRAKECOMMANDOPENCONFIRMED, 'bypass actif : confirmation = image de BrakeCmd');
END_TEST

TEST 'Comportement actuel : fermeture immediate sans attendre DelayMotorDecel (TonDecel jamais cable)'
    (* A VERIFIER intentionnellement : DelayMotorDecel/TonDecel sont declares et documentes
       ("Delai deceleration avant collage frein") mais TonDecel.IN est TOUJOURS force a FALSE
       dans FB_Brake.st (§1/§3) -- aucune temporisation n est reellement appliquee avant que le
       frein ne colle. Ce test documente le comportement REEL actuel (immediat), pas une exigence
       validee -- a confirmer avec l utilisateur si une temporisation etait pourtant voulue. *)
    fb(ENABLE := TRUE, RESET := FALSE, MOVEMENTREQUESTED := TRUE,
       CONTACTORFEEDBACK := FALSE, BYPASSCONTACTORCHECK := TRUE,
       DELAYCONTACTCLOSE := T#100MS, DELAYMAGNETISE := T#300MS,
       DELAYMOTORDECEL := T#500MS, FEEDBACKTIMEOUT := T#1S);
    ADVANCE_TIME(401000000);
    fb(ENABLE := TRUE, RESET := FALSE, MOVEMENTREQUESTED := TRUE,
       CONTACTORFEEDBACK := FALSE, BYPASSCONTACTORCHECK := TRUE,
       DELAYCONTACTCLOSE := T#100MS, DELAYMAGNETISE := T#300MS,
       DELAYMOTORDECEL := T#500MS, FEEDBACKTIMEOUT := T#1S);
    ASSERT_TRUE(fb.BRAKECMD, 'precondition : frein ouvert');

    (* mouvement arrete : meme scan, frein colle instantanement -- DelayMotorDecel (500ms) ignore *)
    ADVANCE_TIME(10000000);
    fb(ENABLE := TRUE, RESET := FALSE, MOVEMENTREQUESTED := FALSE,
       CONTACTORFEEDBACK := FALSE, BYPASSCONTACTORCHECK := TRUE,
       DELAYCONTACTCLOSE := T#100MS, DELAYMAGNETISE := T#300MS,
       DELAYMOTORDECEL := T#500MS, FEEDBACKTIMEOUT := T#1S);
    ASSERT_FALSE(fb.BRAKECMD, 'MovementRequested retombe : frein colle DES CE SCAN, aucun delai observe');
    ASSERT_TRUE(fb.READY, 'FB reste Ready');
END_TEST

TEST 'Double verification contacteur : StuckClosed si le retour ne confirme jamais l ouverture'
    fb(ENABLE := TRUE, RESET := FALSE, MOVEMENTREQUESTED := TRUE,
       CONTACTORFEEDBACK := FALSE, BYPASSCONTACTORCHECK := FALSE,
       DELAYCONTACTCLOSE := T#100MS, DELAYMAGNETISE := T#300MS,
       DELAYMOTORDECEL := T#500MS, FEEDBACKTIMEOUT := T#1S);
    ADVANCE_TIME(401000000);
    fb(ENABLE := TRUE, RESET := FALSE, MOVEMENTREQUESTED := TRUE,
       CONTACTORFEEDBACK := FALSE, BYPASSCONTACTORCHECK := FALSE,
       DELAYCONTACTCLOSE := T#100MS, DELAYMAGNETISE := T#300MS,
       DELAYMOTORDECEL := T#500MS, FEEDBACKTIMEOUT := T#1S);
    ASSERT_TRUE(fb.BRAKECMD, 'magnetisation acquise : commande ouverture emise (ContactorFeedback ne confirme pas encore)');

    (* 1s de plus (FeedbackTimeout) : le retour n a jamais confirme -> defaut *)
    ADVANCE_TIME(1000000000);
    fb(ENABLE := TRUE, RESET := FALSE, MOVEMENTREQUESTED := TRUE,
       CONTACTORFEEDBACK := FALSE, BYPASSCONTACTORCHECK := FALSE,
       DELAYCONTACTCLOSE := T#100MS, DELAYMAGNETISE := T#300MS,
       DELAYMOTORDECEL := T#500MS, FEEDBACKTIMEOUT := T#1S);
    ASSERT_TRUE(fb.CONTACTORCHECK.STUCKCLOSED, 'commande ouverture emise mais jamais confirmee -> StuckClosed');
    ASSERT_TRUE(fb.FAULT.ERROR, 'defaut visible sur Fault.Error');
    ASSERT_TRUE(fb.FAULT.LATCHED, 'defaut latche');
    ASSERT_EQ(fb.FAULT.ERRORID, 16#0001, 'bit0 : incoherence retour contacteur');
    ASSERT_FALSE(fb.BRAKECMD, 'sortie sure sur defaut : BrakeCmd force a FALSE malgre la sequence terminee');
END_TEST

TEST 'Reset n acquitte le defaut contacteur que si la cause (retour) a reellement disparu'
    fb(ENABLE := TRUE, RESET := FALSE, MOVEMENTREQUESTED := TRUE,
       CONTACTORFEEDBACK := FALSE, BYPASSCONTACTORCHECK := FALSE,
       DELAYCONTACTCLOSE := T#100MS, DELAYMAGNETISE := T#300MS,
       DELAYMOTORDECEL := T#500MS, FEEDBACKTIMEOUT := T#1S);
    ADVANCE_TIME(401000000);
    fb(ENABLE := TRUE, RESET := FALSE, MOVEMENTREQUESTED := TRUE,
       CONTACTORFEEDBACK := FALSE, BYPASSCONTACTORCHECK := FALSE,
       DELAYCONTACTCLOSE := T#100MS, DELAYMAGNETISE := T#300MS,
       DELAYMOTORDECEL := T#500MS, FEEDBACKTIMEOUT := T#1S);
    ADVANCE_TIME(1000000000);
    fb(ENABLE := TRUE, RESET := FALSE, MOVEMENTREQUESTED := TRUE,
       CONTACTORFEEDBACK := FALSE, BYPASSCONTACTORCHECK := FALSE,
       DELAYCONTACTCLOSE := T#100MS, DELAYMAGNETISE := T#300MS,
       DELAYMOTORDECEL := T#500MS, FEEDBACKTIMEOUT := T#1S);
    ASSERT_TRUE(fb.FAULT.ERROR, 'precondition : defaut StuckClosed actif');

    (* la cause disparait (le retour confirme enfin), mais SANS Reset : le defaut reste affiche *)
    ADVANCE_TIME(10000000);
    fb(ENABLE := TRUE, RESET := FALSE, MOVEMENTREQUESTED := TRUE,
       CONTACTORFEEDBACK := TRUE, BYPASSCONTACTORCHECK := FALSE,
       DELAYCONTACTCLOSE := T#100MS, DELAYMAGNETISE := T#300MS,
       DELAYMOTORDECEL := T#500MS, FEEDBACKTIMEOUT := T#1S);
    ASSERT_TRUE(fb.FAULT.LATCHED, 'cause disparue mais pas acquittee : le latch reste actif');

    (* front Reset, cause deja disparue : acquitte *)
    ADVANCE_TIME(10000000);
    fb(ENABLE := TRUE, RESET := TRUE, MOVEMENTREQUESTED := TRUE,
       CONTACTORFEEDBACK := TRUE, BYPASSCONTACTORCHECK := FALSE,
       DELAYCONTACTCLOSE := T#100MS, DELAYMAGNETISE := T#300MS,
       DELAYMOTORDECEL := T#500MS, FEEDBACKTIMEOUT := T#1S);
    ASSERT_FALSE(fb.FAULT.ERROR, 'Reset avec cause disparue (retour coherent) : defaut live acquitte');
    ASSERT_FALSE(fb.FAULT.LATCHED, 'Reset avec cause disparue : latch acquitte');
    ASSERT_TRUE(fb.BRAKECMD, 'plus de defaut : frein a nouveau relache (mouvement toujours demande)');
END_TEST

(* ---- FB_CycleTime_test.st ---- *)
SETUP
VAR
    fb : FB_CYCLETIME;
END_VAR
END_SETUP

TEST 'Premier cycle retourne la valeur de secours (pas de dt mesurable)'
    fb(DEFAULTVALUES := 0.004);
    ASSERT_NEAR(fb.CYCLETIMES, 0.004, 0.0001, 'premier appel : aucun dt reel disponible, DefaultValueS renvoye tel quel');
END_TEST

TEST 'Cycle suivant calcule le dt reel ecoule (ms->s)'
    fb(DEFAULTVALUES := 0.004);
    ADVANCE_TIME(10000000);
    fb(DEFAULTVALUES := 0.004);
    ASSERT_NEAR(fb.CYCLETIMES, 0.01, 0.0001, '10ms ecoulees entre les 2 appels -> 0.01s calcule (pas la valeur de secours)');

    ADVANCE_TIME(25000000);
    fb(DEFAULTVALUES := 0.004);
    ASSERT_NEAR(fb.CYCLETIMES, 0.025, 0.0001, 'dt variable d un cycle a l autre correctement mesure (25ms)');

    ADVANCE_TIME(1000000000);
    fb(DEFAULTVALUES := 0.004);
    ASSERT_NEAR(fb.CYCLETIMES, 1.0, 0.0001, 'borne haute INCLUSE : dt = 1000ms = CST_MaxCycleDeltaMs -> dt reel publie (pas secours)');
END_TEST

TEST 'Delta nul (deux appels sans avance horloge) : borne basse -> valeur de secours'
    fb(DEFAULTVALUES := 0.004);
    ADVANCE_TIME(10000000);
    fb(DEFAULTVALUES := 0.004);
    fb(DEFAULTVALUES := 0.004);
    ASSERT_NEAR(fb.CYCLETIMES, 0.004, 0.0001, 'dt = 0 : anti-zero conserve, DefaultValueS publie');
END_TEST

TEST 'Delta aberrant > plafond (5s, simule rebouclage TIME() / reprise) : borne haute -> secours, non latche'
    fb(DEFAULTVALUES := 0.004);
    ADVANCE_TIME(5000000000);
    fb(DEFAULTVALUES := 0.004);
    ASSERT_NEAR(fb.CYCLETIMES, 0.004, 0.0001, 'dt > CST_MaxCycleDeltaMs : artefact non propage, DefaultValueS publie');

    ADVANCE_TIME(1001000000);
    fb(DEFAULTVALUES := 0.004);
    ASSERT_NEAR(fb.CYCLETIMES, 0.004, 0.0001, 'borne haute EXCLUE : dt = 1001ms (juste au-dessus du plafond) -> DefaultValueS');

    ADVANCE_TIME(10000000);
    fb(DEFAULTVALUES := 0.004);
    ASSERT_NEAR(fb.CYCLETIMES, 0.01, 0.0001, 'scan suivant a dt nominal : le dt reel est de nouveau publie (secours non latche)');
END_TEST

(* ---- FB_FaultCore_test.st ---- *)
(* =======================================================================
   🧪 test_fb_faultcore.st — Socle FB_FaultCore (TC-P03-008..013)
   ───────────────────────────────────────────────────────────────
   Lot : T174 (P0 — test_fb_fbstatus.st vise un FB supprimé au commit
   51fccce6 ; CE fichier le remplace contre FB_FaultCore.st actuel.
   Fiche : DOC/AF/AF_Partie-03_Contrats_Composants/FB_FaultCore_v1.0.md §2.
   Conventions : 1 appel fb() = 1 scan ; ADVANCE_TIME(10000000) entre les
   scans pour les fronts R_TRIG ; hex décrit en décimal (bit 0 = 1, bit 15 = 32768).
   ======================================================================= *)

SETUP
VAR
    fb : FB_FAULTCORE;
END_VAR
END_SETUP

(* ── Remise à zéro commune : pulse Enable+Reset, puis Reset retombé ── *)

TEST 'TC-P03-011 Reset sans historique de defaut : aucun effet parasite'
    (* Remise à zéro avec un front Reset sur un FB vierge *)
    fb(ENABLE := TRUE, RESET := TRUE);
    ADVANCE_TIME(10000000);
    fb(ENABLE := TRUE, RESET := FALSE);
    ADVANCE_TIME(10000000);
    ASSERT_EQ(fb.FAULT.LATCHEDID, 0, 'Reset sans historique : LatchedId reste 0');
    ASSERT_FALSE(fb.FAULT.LATCHED, 'Reset sans historique : Latched reste FALSE');
    ASSERT_EQ(fb.FAULT.ERRORID, 0, 'Aucune cause active : ErrorId = 0');
    ASSERT_FALSE(fb.FAULT.ERROR, 'Aucune cause active : Error = FALSE');
    ASSERT_TRUE(fb.READY, 'Enable=TRUE -> Ready=TRUE');
END_TEST

TEST 'TC-P03-008 Cumul de 2 causes latchees apparues a des instants differents, un seul Reset les acquitte ensemble'
    (* Remise a zero *)
    fb(ENABLE := TRUE, RESET := TRUE);
    ADVANCE_TIME(10000000);
    fb(ENABLE := TRUE, RESET := FALSE);

    (* Cause 2 latchee apparait -> bit 2 (4) latche ; causes inactives entre scans *)
    fb.CAUSES[2].ACTIVE := TRUE;
    fb.CAUSES[2].LATCHING := TRUE;
    fb(ENABLE := TRUE, RESET := FALSE);
    ASSERT_EQ(fb.FAULT.LATCHEDID, 4, 'Cause 2 latchee -> LatchedId = bit 2 (4)');
    ASSERT_TRUE(fb.FAULT.LATCHED, 'Latch arme');

    (* La cause 2 disparait -> le bit latche reste (defaut non acquitte) *)
    fb.CAUSES[2].ACTIVE := FALSE;
    ADVANCE_TIME(10000000);
    fb(ENABLE := TRUE, RESET := FALSE);
    ASSERT_EQ(fb.FAULT.LATCHEDID, 4, 'Cause disparue, bit 2 latche conserve');
    ASSERT_FALSE(fb.FAULT.ERROR, 'Cause 2 inactive : vue LIVE retombee');

    (* Cause 5 latchee apparait a un autre instant -> cumul bits 2 + 5 (4 + 32 = 36) *)
    fb.CAUSES[5].ACTIVE := TRUE;
    fb.CAUSES[5].LATCHING := TRUE;
    fb(ENABLE := TRUE, RESET := FALSE);
    ASSERT_EQ(fb.FAULT.LATCHEDID, 36, 'Cumul bit 2 (4) + bit 5 (32) = 36');
    ASSERT_TRUE(fb.FAULT.ERROR, 'Cause 5 active -> vue LIVE en erreur');

    (* Les 2 causes se relâchent SANS Reset (ré-armement fail-safe : le bit reste tant
       que la cause est active — il faut désactiver AVANT d'asserter le clear) *)
    fb.CAUSES[5].ACTIVE := FALSE;
    ADVANCE_TIME(10000000);
    fb(ENABLE := TRUE, RESET := FALSE);
    ASSERT_EQ(fb.FAULT.LATCHEDID, 36, 'Causes relâchées sans Reset : les 2 latches (36) restent');
    ASSERT_FALSE(fb.FAULT.ERROR, 'Vue LIVE retombée (aucune cause active)');

    (* Un seul front Reset les acquitte ensemble *)
    fb(ENABLE := TRUE, RESET := TRUE);
    ADVANCE_TIME(10000000);
    fb(ENABLE := TRUE, RESET := FALSE);
    ASSERT_EQ(fb.FAULT.LATCHEDID, 0, 'Un seul front Reset acquitte les 2 latches ensemble');
    ASSERT_FALSE(fb.FAULT.LATCHED, 'Plus aucun latch apres Reset');

    (* Nettoyage causes pour la suite *)
    fb.CAUSES[2].ACTIVE := FALSE;
    fb.CAUSES[2].LATCHING := FALSE;
    fb.CAUSES[5].ACTIVE := FALSE;
    fb.CAUSES[5].LATCHING := FALSE;
    fb(ENABLE := TRUE, RESET := FALSE);
END_TEST

TEST 'TC-P03-009 Cause live + cause latchee simultanees : live retombe seule, latchee reste jusqu au Reset'
    (* Remise a zero *)
    fb(ENABLE := TRUE, RESET := TRUE);
    ADVANCE_TIME(10000000);
    fb(ENABLE := TRUE, RESET := FALSE);

    (* Cause 1 live + cause 3 latchee simultanees (aligne sur la fiche TC-P03-009) *)
    fb.CAUSES[1].ACTIVE := TRUE;
    fb.CAUSES[1].LATCHING := FALSE;
    fb.CAUSES[3].ACTIVE := TRUE;
    fb.CAUSES[3].LATCHING := TRUE;
    fb(ENABLE := TRUE, RESET := FALSE);
    ASSERT_EQ(fb.FAULT.ERRORID, 10, 'ErrorId LIVE = bit 1 (2) + bit 3 (8) = 10');
    ASSERT_TRUE(fb.FAULT.ERROR, 'Deux causes actives -> Error=TRUE');
    ASSERT_EQ(fb.FAULT.LATCHEDID, 8, 'LatchedId = bit 3 (8) seul (cause 1 non latchee)');

    (* La cause live retombe seule : elle quitte ErrorId (bit 3 reste : cause 3 ENCORE active) *)
    fb.CAUSES[1].ACTIVE := FALSE;
    ADVANCE_TIME(10000000);
    fb(ENABLE := TRUE, RESET := FALSE);
    ASSERT_EQ(fb.FAULT.ERRORID, 8, 'Cause 1 inactive -> ErrorId = bit 3 seul (cause 3 encore active)');
    ASSERT_TRUE(fb.FAULT.ERROR, 'Cause 3 toujours active -> Error=TRUE');
    ASSERT_EQ(fb.FAULT.LATCHEDID, 8, 'Latche conservee apres retombee de la live');

    (* La latchee se relache elle aussi SANS Reset : latches conservees (fail-safe),
       MAIS ErrorId retombe (plus aucune cause active) *)
    fb.CAUSES[3].ACTIVE := FALSE;
    ADVANCE_TIME(10000000);
    fb(ENABLE := TRUE, RESET := FALSE);
    ASSERT_EQ(fb.FAULT.ERRORID, 0, 'Cause 3 inactive -> ErrorId = 0 sans Reset');
    ASSERT_EQ(fb.FAULT.LATCHEDID, 8, 'Latche conservee apres disparition de la cause');

    (* Front Reset : la latchee est acquitte *)
    fb(ENABLE := TRUE, RESET := TRUE);
    ADVANCE_TIME(10000000);
    fb(ENABLE := TRUE, RESET := FALSE);
    ASSERT_EQ(fb.FAULT.LATCHEDID, 0, 'Reset front efface la latchee');

    (* Nettoyage *)
    fb.CAUSES[1].ACTIVE := FALSE;
    fb.CAUSES[1].LATCHING := FALSE;
    fb(ENABLE := TRUE, RESET := FALSE);
END_TEST

TEST 'TC-P03-010 Bornes de la liste Causes : bit 0 et bit 15 correctement mappes (pas d off-by-one)'
    (* Remise a zero *)
    fb(ENABLE := TRUE, RESET := TRUE);
    ADVANCE_TIME(10000000);
    fb(ENABLE := TRUE, RESET := FALSE);

    (* Causes[0] et Causes[15] latchees et actives *)
    fb.CAUSES[0].ACTIVE := TRUE;
    fb.CAUSES[0].LATCHING := TRUE;
    fb.CAUSES[15].ACTIVE := TRUE;
    fb.CAUSES[15].LATCHING := TRUE;
    fb(ENABLE := TRUE, RESET := FALSE);
    ASSERT_EQ(fb.FAULT.LATCHEDID, 32769, 'Bit 0 (1) + bit 15 (32768) = 32769, pas d off-by-one');
    ASSERT_EQ(fb.FAULT.ERRORID, 32769, 'Vue LIVE identique : SHL(1, i) aux bornes');

    (* Les 2 causes se relachent SANS Reset : les latches (32769) restent (fail-safe) *)
    fb.CAUSES[0].ACTIVE := FALSE;
    fb.CAUSES[15].ACTIVE := FALSE;
    ADVANCE_TIME(10000000);
    fb(ENABLE := TRUE, RESET := FALSE);
    ASSERT_EQ(fb.FAULT.LATCHEDID, 32769, 'Causes relachees sans Reset : latches conservees');
    ASSERT_EQ(fb.FAULT.ERRORID, 0, 'Vue LIVE retombee : ErrorId = 0 sans Reset');

    (* Front Reset *)
    fb(ENABLE := TRUE, RESET := TRUE);
    ADVANCE_TIME(10000000);
    fb(ENABLE := TRUE, RESET := FALSE);
    ASSERT_EQ(fb.FAULT.LATCHEDID, 0, 'Reset aux bornes : rien ne persiste');

    (* Nettoyage *)
    fb.CAUSES[0].ACTIVE := FALSE;
    fb.CAUSES[0].LATCHING := FALSE;
    fb.CAUSES[15].ACTIVE := FALSE;
    fb.CAUSES[15].LATCHING := FALSE;
    fb(ENABLE := TRUE, RESET := FALSE);
END_TEST

TEST 'TC-P03-012 Reset maintenu niveau haut : pas d acquittement silencieux, cause reaparue re-arme (faille T148 non applicable)'
    (* Remise a zero *)
    fb(ENABLE := TRUE, RESET := TRUE);
    ADVANCE_TIME(10000000);
    fb(ENABLE := TRUE, RESET := FALSE);

    (* Cause 0 latchee -> LatchedId = 1 *)
    fb.CAUSES[0].ACTIVE := TRUE;
    fb.CAUSES[0].LATCHING := TRUE;
    fb(ENABLE := TRUE, RESET := FALSE);
    ASSERT_EQ(fb.FAULT.LATCHEDID, 1, 'Cause latchee -> bit 0');

    (* Reset passe TRUE (nouveau front) pendant que la cause est inactive : clear legitime *)
    fb.CAUSES[0].ACTIVE := FALSE;
    ADVANCE_TIME(10000000);
    fb(ENABLE := TRUE, RESET := TRUE);
    ADVANCE_TIME(10000000);
    fb(ENABLE := TRUE, RESET := TRUE);
    ASSERT_EQ(fb.FAULT.LATCHEDID, 0, 'Front Reset (cause inactive) : latches effaces');

    (* Reset MAINTENU (T#TRUE, aucun nouveau front) : la cause reapparait -> re-armement fail-safe *)
    fb.CAUSES[0].ACTIVE := TRUE;
    ADVANCE_TIME(10000000);
    fb(ENABLE := TRUE, RESET := TRUE);
    ASSERT_EQ(fb.FAULT.LATCHEDID, 1, 'Cause reapparue Active AND Latching sous Reset maintenu : re-arme (pas d acquittement silencieux)');

    (* Cause redisparait, Reset TOUJOURS maintenu : aucun nouveau front -> le bit re-arme n est PAS efface *)
    fb.CAUSES[0].ACTIVE := FALSE;
    ADVANCE_TIME(10000000);
    fb(ENABLE := TRUE, RESET := TRUE);
    ASSERT_EQ(fb.FAULT.LATCHEDID, 1, 'R_TRIG sans nouveau front : le clear ne s applique pas (faille T148 non applicable)');

    (* Reset relache puis re-pulse : acquittement effectif *)
    ADVANCE_TIME(10000000);
    fb(ENABLE := TRUE, RESET := FALSE);
    ADVANCE_TIME(10000000);
    fb(ENABLE := TRUE, RESET := TRUE);
    ADVANCE_TIME(10000000);
    fb(ENABLE := TRUE, RESET := FALSE);
    ASSERT_EQ(fb.FAULT.LATCHEDID, 0, 'Nouveau front Reset apres relachement : acquittement effectif');

    (* Nettoyage *)
    fb.CAUSES[0].ACTIVE := FALSE;
    fb.CAUSES[0].LATCHING := FALSE;
    fb(ENABLE := TRUE, RESET := FALSE);
END_TEST

TEST 'TC-P03-013 Enable=FALSE : vue LIVE masquee mais vue LATCHEE reste publiee (pas d effacement silencieux OFF->ON)'
    (* Remise a zero *)
    fb(ENABLE := TRUE, RESET := TRUE);
    ADVANCE_TIME(10000000);
    fb(ENABLE := TRUE, RESET := FALSE);

    (* Cause latchee apparait et latche *)
    fb.CAUSES[1].ACTIVE := TRUE;
    fb.CAUSES[1].LATCHING := TRUE;
    fb(ENABLE := TRUE, RESET := FALSE);
    ASSERT_EQ(fb.FAULT.LATCHEDID, 2, 'Cause 1 latchee -> bit 1 (2)');

    (* Enable=FALSE : LIVE masquee, LATCHED conserve *)
    fb(ENABLE := FALSE, RESET := FALSE);
    ADVANCE_TIME(10000000);
    fb(ENABLE := FALSE, RESET := FALSE);
    ASSERT_EQ(fb.FAULT.ERRORID, 0, 'Enable=FALSE : vue LIVE non evaluee -> ErrorId=0');
    ASSERT_FALSE(fb.FAULT.ERROR, 'Enable=FALSE : Error=FALSE');
    ASSERT_EQ(fb.FAULT.LATCHEDID, 2, 'Enable=FALSE : LatchedId CONSERVE (pas d effacement silencieux)');
    ASSERT_TRUE(fb.FAULT.LATCHED, 'Latche toujours publiee meme FB desactive');

    (* Retour Enable=TRUE SANS Reset : le latch reste (bascule OFF->ON n efface rien) *)
    fb(ENABLE := TRUE, RESET := FALSE);
    ADVANCE_TIME(10000000);
    fb(ENABLE := TRUE, RESET := FALSE);
    ASSERT_EQ(fb.FAULT.LATCHEDID, 2, 'Re-Enable sans Reset : latch conserve (bascule OFF->ON n efface rien)');

    (* Reset aussi effectif avec Enable=FALSE (std §9 : jamais conditionne) *)
    fb(ENABLE := FALSE, RESET := TRUE);
    ADVANCE_TIME(10000000);
    fb(ENABLE := FALSE, RESET := FALSE);
    ASSERT_EQ(fb.FAULT.LATCHEDID, 0, 'Reset front agit meme Enable=FALSE');

    (* Nettoyage *)
    fb.CAUSES[1].ACTIVE := FALSE;
    fb.CAUSES[1].LATCHING := FALSE;
    fb(ENABLE := TRUE, RESET := FALSE);
END_TEST

(* =======================================================================
   Règles générales du socle Cause/Ack (AF_Partie-03 §4) — TC-P03-003/004/005.
   Le socle FB_FaultCore illustre ces règles transverses : pas de redémarrage
   auto après Ack (003), pas de SafeStop/StartStop hors mouvement (004),
   encapsulation stricte (005).
   ======================================================================= *)

TEST 'TC-P03-003 Pas de redemarrage auto apres Ack : Reset retourne Ready, un nouvel ordre explicite est requis'
    (* Remise a zero *)
    fb(ENABLE := TRUE, RESET := TRUE);
    ADVANCE_TIME(10000000);
    fb(ENABLE := TRUE, RESET := FALSE);

    (* Cause 0 latchee -> LatchedId = 1 *)
    fb.CAUSES[0].ACTIVE := TRUE;
    fb.CAUSES[0].LATCHING := TRUE;
    fb(ENABLE := TRUE, RESET := FALSE);
    ASSERT_EQ(fb.FAULT.LATCHEDID, 1, 'Cause latchee -> bit 0');

    (* Front Reset (Ack) : efface le latch, retour Ready *)
    fb.CAUSES[0].ACTIVE := FALSE;
    ADVANCE_TIME(10000000);
    fb(ENABLE := TRUE, RESET := TRUE);
    ADVANCE_TIME(10000000);
    fb(ENABLE := TRUE, RESET := FALSE);
    ASSERT_EQ(fb.FAULT.LATCHEDID, 0, 'Ack (Reset) efface le latch');
    ASSERT_TRUE(fb.READY, 'Apres Ack, le FB est Ready');

    (* Pas de redemarrage auto : sans nouvelle cause, le latch reste 0 sur plusieurs scans *)
    ADVANCE_TIME(10000000);
    fb(ENABLE := TRUE, RESET := FALSE);
    ASSERT_EQ(fb.FAULT.LATCHEDID, 0, 'Aucun re-armement auto apres Ack (scan 1)');
    ADVANCE_TIME(10000000);
    fb(ENABLE := TRUE, RESET := FALSE);
    ASSERT_EQ(fb.FAULT.LATCHEDID, 0, 'Aucun re-armement auto apres Ack (scan 2)');

    (* Un nouvel ordre explicite (nouvelle cause Active AND Latching) re-arme *)
    fb.CAUSES[0].ACTIVE := TRUE;
    fb(ENABLE := TRUE, RESET := FALSE);
    ASSERT_EQ(fb.FAULT.LATCHEDID, 1, 'Nouvelle cause explicite -> re-armement (pas auto)');

    (* Nettoyage *)
    fb.CAUSES[0].ACTIVE := FALSE;
    fb.CAUSES[0].LATCHING := FALSE;
    fb(ENABLE := TRUE, RESET := FALSE);
END_TEST

TEST 'TC-P03-004 Pas de SafeStop/StartStop hors mouvement (invariant structurel)'
    (* 💻 AUTO — invariant structurel documenté, pas un comportement runtime.
       Règle AF_Partie-03 §3 : SafeStop/StartStop ne sont autorisés QUE sur un FB
       de mouvement. Le socle FB_FaultCore (brique technique transverse) n'expose
       NI SafeStop NI StartStop dans son interface : VAR_INPUT = Enable/Reset/Causes,
       VAR_OUTPUT = Ready/Fault. Aucun SafeStop/StartStop n'est donc possible ici.
       Vérifié structurellement par l'interface déclarée (pas de port de mouvement). *)
    fb(ENABLE := TRUE, RESET := FALSE);
    ASSERT_TRUE(fb.READY, 'socle actif -> Ready=TRUE (aucun port de mouvement a tester)');
END_TEST

TEST 'TC-P03-005 Encapsulation stricte : echanges via interfaces/DUTs publics uniquement (invariant structurel)'
    (* 💻 AUTO — invariant structurel documenté, pas un comportement runtime.
       Règle AF_Partie-03 §2 : les variables internes sont privées, les échanges
       passent uniquement par interfaces et DUT publics. FB_FaultCore n'expose que
       ses VAR_INPUT (Enable/Reset/Causes) et VAR_OUTPUT (Ready/Fault) ; ses internes
       (ResetEdge, Latch[], i) sont privés. Vérifié par encapsulation_check.py
       (aucune écriture externe non déclarée, aucun accès GVL direct). *)
    fb(ENABLE := TRUE, RESET := FALSE);
    ASSERT_TRUE(fb.READY, 'socle accessible par son interface publique uniquement');
END_TEST

(* ---- FB_Filter_test.st ---- *)
SETUP
VAR
    fb : FB_FILTER;
END_VAR
END_SETUP

TEST 'Pass-through si TimeConst=0 (pas de lissage)'
    fb(VALUEIN := 10.0, TIMECONST := T#0MS, CYCLETIMES := 0.1);
    ASSERT_NEAR(fb.VALUEOUT, 10.0, 0.001, 'TimeConst=0 -> recopie directe de ValueIn');
END_TEST

TEST 'Pass-through si CycleTimeS=0 (temps de cycle invalide)'
    fb(VALUEIN := 10.0, TIMECONST := T#200MS, CYCLETIMES := 0.0);
    ASSERT_NEAR(fb.VALUEOUT, 10.0, 0.001, 'CycleTimeS=0 -> recopie directe de ValueIn (garde-fou division par zero)');
END_TEST

TEST 'Reponse PT1 : convergence progressive vers un echelon, pas instantanee'
    (* TimeConst=100ms, CycleTimeS=100ms -> Alpha = 0.1/(0.1+0.1) = 0.5 *)
    fb(VALUEIN := 10.0, TIMECONST := T#100MS, CYCLETIMES := 0.1);
    ASSERT_NEAR(fb.VALUEOUT, 5.0, 0.001, 'scan 1 : ValueOut = 0.5*10 + 0.5*0 = 5.0 (pas de saut brutal a 10)');

    fb(VALUEIN := 10.0, TIMECONST := T#100MS, CYCLETIMES := 0.1);
    ASSERT_NEAR(fb.VALUEOUT, 7.5, 0.001, 'scan 2 : ValueOut = 0.5*10 + 0.5*5 = 7.5 (memoire du scan precedent)');

    fb(VALUEIN := 10.0, TIMECONST := T#100MS, CYCLETIMES := 0.1);
    ASSERT_NEAR(fb.VALUEOUT, 8.75, 0.001, 'scan 3 : ValueOut = 0.5*10 + 0.5*7.5 = 8.75 (convergence exponentielle vers 10)');
END_TEST

(* ---- FB_Ramp_test.st ---- *)
SETUP
VAR
    fb : FB_RAMP;
END_VAR
END_SETUP

TEST 'Accel : consigne progresse par pas de AccelRate*CycleTimeS vers la cible'
    fb(TARGET := 100.0, ACCELRATE := 50.0, DECELRATE := 200.0, CYCLETIMES := 0.1);
    ASSERT_NEAR(fb.CURRENT, 5.0, 0.001, 'pas 1 : 0 -> 5.0 (50%/s * 0.1s), s eloigne de zero donc AccelRate');

    fb(TARGET := 100.0, ACCELRATE := 50.0, DECELRATE := 200.0, CYCLETIMES := 0.1);
    ASSERT_NEAR(fb.CURRENT, 10.0, 0.001, 'pas 2 : 5.0 -> 10.0, meme taux tant que la cible n est pas atteinte');
END_TEST

TEST 'Decel : retour vers zero utilise DecelRate (taux different d Accel)'
    (* monte a 40% avec Accel *)
    fb(TARGET := 40.0, ACCELRATE := 50.0, DECELRATE := 10.0, CYCLETIMES := 0.1);
    ASSERT_NEAR(fb.CURRENT, 5.0, 0.001, 'montee : AccelRate (50%/s)');
    fb(TARGET := 40.0, ACCELRATE := 50.0, DECELRATE := 10.0, CYCLETIMES := 0.1);
    ASSERT_NEAR(fb.CURRENT, 10.0, 0.001, 'montee : toujours AccelRate, cible pas encore atteinte');

    (* cible ramenee a 0 : retour vers zero -> DecelRate, taux bien plus faible ici *)
    fb(TARGET := 0.0, ACCELRATE := 50.0, DECELRATE := 10.0, CYCLETIMES := 0.1);
    ASSERT_NEAR(fb.CURRENT, 9.0, 0.001, 'retour vers zero : DecelRate (10%/s), pas de 1.0 seulement -- pas AccelRate');
END_TEST

TEST 'Atteinte de la cible : la rampe s arrete pile dessus, pas de depassement'
    fb(TARGET := 3.0, ACCELRATE := 50.0, DECELRATE := 200.0, CYCLETIMES := 0.1);
    ASSERT_NEAR(fb.CURRENT, 3.0, 0.001, 'le pas (5.0) depasserait la cible (3.0) : clampe exactement dessus, pas de depassement');

    fb(TARGET := 3.0, ACCELRATE := 50.0, DECELRATE := 200.0, CYCLETIMES := 0.1);
    ASSERT_NEAR(fb.CURRENT, 3.0, 0.001, 'cible deja atteinte : reste stable, aucune oscillation autour de la cible');
END_TEST

TEST 'Garde-fou : une valeur Current deja hors plage (etat corrompu) reste bornee a +/-100'
    (* Simule un etat interne deja corrompu au-dela de la plage normalisee -- le FB doit se
       proteger lui-meme, pas seulement empecher d y entrer *)
    fb(TARGET := 500.0, ACCELRATE := 1000.0, DECELRATE := 1000.0, CYCLETIMES := 1.0);
    ASSERT_NEAR(fb.CURRENT, 100.0, 0.001, 'Target hors plage (500) et grand pas (1000%/s) : Current ne depasse jamais +100');
END_TEST
